// TIA Portal V21 export
// export: Created 2026-10-14T03:11:20.5445002Z, ExportSetting WithDefaults, DisplayName Totally Integrated Automation Portal, DisplayVersion V21, DisplayName STEP 7 Professional, DisplayVersion V21, DisplayName STEP 7 Safety, DisplayVersion V21, DisplayName Tech WebApplication, DisplayVersion V21, DisplayName WinCC Basic/Comfort/Advanced, DisplayVersion V21, DisplayName WinCC Unified, DisplayVersion V21
TagTable "_RUN"
  RUN_DB_resetAll : Bool  (HMI_Connection_1, 100 ms)
  RUN_DB_resetPID : Bool  (HMI_Connection_1, 100 ms)
  RUN_DB_resetPvSim : Bool  (HMI_Connection_1, 100 ms)
  RUN_DB_resetAccErr : Bool  (HMI_Connection_1, 1 s)
  RUN_DB_setpoint : Real  (HMI_Connection_1, 1 s)
